Fanuc KAREL source: kt00236.KL

-- PROVISIONAL review KL for V1013-1; original PC SHA256 dd37ba914b7403179f3774f675f5d2d54d368150a58bf7033b8df9131daac811
-- Incomplete behavior may be omitted. Consult companion uncertainty JSON. Do not deploy.
PROGRAM KT00236
%NOLOCKGROUP
VAR
  I1 : INTEGER
  I2 : INTEGER
  OUT : INTEGER
BEGIN
  -- UNRESOLVED_PC offsets 5-16; opcodes 2E,23
  -- UNRESOLVED_PC offsets 21-32; opcodes 2E,23
  -- UNRESOLVED_PC offsets 37-48; opcodes 2E,23
  -- UNRESOLVED_PC offsets 53-64; opcodes 2E,23
  -- UNRESOLVED_PC offsets 69-88; opcodes 21,21,47,23
  -- UNRESOLVED_PC offsets 93-97; opcodes 7F
END KT00236
